{region 'Documentation'}
(*!
<summary>Checks inequality with the forbidden BYTE value.</summary>
*)
{endregion}
FUNCTION_BLOCK AssertNotEqual_Byte EXTENDS AssertionBase
VAR_INPUT
    IN : BYTE; //! Actual value checked or observed by this Assertion.
    Expected : BYTE; //! Value that must differ from IN under this Assertion's comparison rules.
END_VAR

SUPER^();

{region 'Documentation'}
(*!
<summary>Check inequality with the forbidden BYTE value.</summary>
*)
{endregion}
METHOD PROTECTED Assert
VAR
    Message : STRING(GVL_Constants.MessageLength);
    ExpectedText : STRING(GVL_Constants.AssertionValueLength);
    ActualText : STRING(GVL_Constants.AssertionValueLength);
END_VAR
VAR CONSTANT
    HexDigitCount : USINT := 2;
END_VAR
IF NOT EvaluationActive THEN
    RETURN;
END_IF;

IF Result = E_Result.Error THEN
    RETURN;
END_IF;

IF Result = E_Result.Failed THEN
    RETURN;
END_IF;

IF IN = Expected THEN
    ExpectedText := CreateAssertionTextValue_Hex(Value := BYTE_TO_LWORD(Expected),
        DigitCount := HexDigitCount);
    ActualText := CreateAssertionTextValue_Hex(Value := BYTE_TO_LWORD(IN),
        DigitCount := HexDigitCount);
    Message := CONCAT('Assertion failed: values are equal but should differ. NotExpected = ',
        ExpectedText);
    Message := CONCAT(Message, ', Actual = ');
    Message := CONCAT(Message, ActualText);
    Message := CONCAT(Message, '.');
    Fail(Message := Message);
    RETURN;
END_IF;

Pass();
END_METHOD

END_FUNCTION_BLOCK

(* stored: Version 1.1.0.1
   POU AssertNotEqual_Byte: Id {d651380b-a6c1-4cb6-966d-c59f59bbe624}, SpecialFunc None
   Folder Internal: Id {d211744a-e9be-4760-a996-2a29a7abbf38}
   Method Assert: Id {732eafe1-b990-4664-be15-16630abfb41e} *)
